Fanuc KAREL source: KA00141.KL

PROGRAM KA00141
%NOLOCKGROUP
VAR
  SRC: ARRAY[2] OF SHORT
  DST: VECTOR
BEGIN
  SRC[1] = 2
  DST = SRC[1]
END KA00141
